FUNCTION_BLOCK StubPart IMPLEMENTS I_XtsPart
VAR_INPUT
END_VAR
VAR_OUTPUT
END_VAR
VAR
END_VAR

{warning 'Add property implementation'}
PROPERTY HasError : BOOL
GET
END_GET
END_PROPERTY

{warning 'Add property implementation'}
PROPERTY Initialised : BOOL
GET
END_GET
END_PROPERTY

{warning 'Add property implementation'}
PROPERTY PartStatus : Xts_Library.XtsPartStatus
GET
END_GET
END_PROPERTY

{warning 'Add method implementation '}
METHOD ResetPart : BOOL
END_METHOD

{warning 'Add method implementation '}
METHOD SetPartOriginTransform : BOOL
VAR_INPUT
	OriginTransform	: Xts_Library.Tc3_XTS_Utility.ST_OriginTransform;
END_VAR
END_METHOD

END_FUNCTION_BLOCK

(* stored: Version 1.1.0.1
   POU StubPart: Id {17764eb3-4e03-4888-b354-67eed1c30915}, SpecialFunc None
   Property HasError: Id {4a26f49f-962b-4fce-ac3a-1eea3e6c74b4}
   Get Get: Id {1910ef9e-c216-41f6-9eb6-a1f3a606f7a4}
   Property Initialised: Id {7449a430-9e1d-4d81-b5d2-ca53e144ce0b}
   Get Get: Id {70a577c7-e31a-41e4-aeb3-913fe1d722cb}
   Property PartStatus: Id {722ab0b3-aa8a-47de-a4f5-1deb35c51a40}
   Get Get: Id {60a133d5-e0ad-4d36-a7bd-fac678a9bfa8}
   Method ResetPart: Id {6ecad392-6345-4f1d-8320-f0009ef7b7f2}
   Method SetPartOriginTransform: Id {0b007cd2-4639-437a-a1e5-de5d60f978b1} *)
